// TIA Portal V19 export
// export: Created 2026-10-16T08:35:17.7165193Z, ExportSetting WithDefaults, DisplayName Totally Integrated Automation Portal, DisplayVersion V19, DisplayName TIA Portal Openness, DisplayVersion V19, DisplayName TIA Portal Version Control Interface, DisplayVersion V19, DisplayName STEP 7 Professional, DisplayVersion V19, DisplayName STEP 7 Safety, DisplayVersion V19, DisplayName WinCC Basic/Comfort/Advanced, DisplayVersion V19, DisplayName WinCC Unified, DisplayVersion V19
TagTable "Default tag table"
  WzorLiczba : Int  (PLC tag ROLL_HMI.Dwell1Seconds, ROLL_PLC, 1 s)
  WzorStan : Bool  (PLC tag ROLL_HMI.Connected, ROLL_PLC, 1 s)
  WzorPrzycisk : Bool  (1 s)
